Staubli VAL3: utCombo.pjx

--- utCombo.pjx ---
Parameters version=s8.8.3Cs9_BS1660 stackSize=5000 millimeterUnit=true
Program file=start.pgx
Program file=stop.pgx
Data file=utCombo.dtx
Type name=utAppearance path=./utAppearance/utAppearance.pjx
Type name=utBorder path=./utBorder/utBorder.pjx
Type name=utCommon path=./utCommon/utCommon.pjx
Type name=utText path=./utText/utText.pjx
Type name=utData path=./utData/utData.pjx

--- utCombo.dtx ---
public utAppearance Appearance
  [0]
    string sBackgroundColour
    string sColour
    bool bVisibility
public utBorder Border
  [0]
    string sBorderColour
    string sBorderStyle
    string sBorderWidth
public utCommon Common
  [0]
    bool bDisabled
    string sValue
    string sID
    string sOption{}
    string sItem
    string sPage
public utText Text
  [0]
    string sFontFamily
    string sFontStyle
    num nFontSize
public utData Data
  [0]
    num nVal
    bool bStatus

--- start.pgx ---
program start()
begin
end

--- stop.pgx ---
program stop()
begin
end
